(* IEC 61131-3 sources: plc-process-lib/src/POUs/Alarm/FB_Alarm, 9 files *)

(* ---- FB_Alarm.decl.st ---- *)
// Назначение: одна тревога по ISA-18.2. Четыре базовых состояния (Normal, ActiveUnack,
//             ActiveAck, RtnUnack) и три наложенных по старшинству OutOfService >
//             SuppressedByDesign > Shelved; приоритет, задержки появления и снятия (FB_Delay),
//             shelve с таймаутом, подавление по условию, вывод из работы. Каждый переход eState
//             увеличивает udiSeq и отправляет событие в GVL_Lib.itfAlarmSink (если приёмник задан).
//             Методы Ack, Shelve, Unshelve только ставят запрос: его выполняет ближайший вызов тела.
//             Модель состояний и повторное оповещение после shelve — сверить с ANSI/ISA-18.2-2016.
// Автор:      kr0nsch
// Версия:     0.1.0
// Документ:   docs/fb/FB_Alarm.md
FUNCTION_BLOCK FB_Alarm IMPLEMENTS I_Alarm
VAR_INPUT
    xIn           : BOOL;            // условие тревоги (до задержек)
    xSuppress     : BOOL;            // подавление по условию (suppressed by design)
    xOutOfService : BOOL;            // вывод из работы (устройство в OutOfService)
    udiId         : UDINT;           // номер тревоги на объекте
    rValue        : REAL;            // значение процесса для события
    stCfg         : ST_AlarmCfg;     // параметры; 16 байт — копирование дешевле ссылки
    itfTime       : I_TimeSource;    // источник времени; 0 — встроенный fbSysTime
END_VAR
VAR_OUTPUT
    eState        : E_AlarmState := E_AlarmState.Normal;   // состояние ISA-18.2
    xActive       : BOOL;            // условие после задержек (независимо от наложенных состояний)
    xUnacked      : BOOL;            // eState = ActiveUnack OR RtnUnack
    xInList       : BOOL;            // ActiveUnack, ActiveAck или RtnUnack — показывать в списке тревог
    xShelved      : BOOL;            // shelve действует (даже если сверху подавление или OutOfService)
    tShelveRemain : TIME;            // остаток shelve; T#0S — shelve нет
    ltLastChange  : LTIME;           // время последнего перехода
    udiSeq        : UDINT;           // +1 на каждый переход eState (переполнение допустимо)
END_VAR
VAR
    fbDelay      : FB_Delay;         // задержки появления (tOnDelay) и снятия (tOffDelay)
    fbSysTime    : FB_SystemTime;    // запасной источник времени
    xAckReq      : BOOL;             // запрос Ack()
    xShelveReq   : BOOL;             // запрос Shelve()
    tShelveReq   : TIME;             // срок из запроса Shelve()
    xUnshelveReq : BOOL;             // запрос Unshelve()
    ltShelveEnd  : LTIME;            // конец действующего shelve
    // --- реализация (сверх контракта 10.1) ---
    ltNow        : LTIME;            // время этого вызова: отметка переходов и событий
    tShelveDur   : TIME;             // срок действующего shelve (после замены T#0S и обрезки)
    ePrioAct     : E_AlarmPriority := E_AlarmPriority.Medium;      // действующий приоритет
    eShelveEnd   : E_AlarmEventReason := E_AlarmEventReason.None;  // как закончился shelve в этом вызове
END_VAR
VAR_TEMP
    itfTimeAct   : I_TimeSource;     // действующий источник этого вызова
END_VAR

(* ---- FB_Alarm.impl.st ---- *)
// 1. Время этого вызова — один раз, для задержек и для отметок событий
IF itfTime <> 0 THEN
    itfTimeAct := itfTime;
ELSE
    itfTimeAct := fbSysTime;
END_IF
ltNow := itfTimeAct.Now();

// 2. Действующий приоритет: значение вне перечисления (мусор persistent-памяти) считается Medium.
//    Строгое перечисление защищает только исходный текст, поэтому проверка — сравнениями
IF stCfg.ePriority = E_AlarmPriority.None OR stCfg.ePriority = E_AlarmPriority.Low
   OR stCfg.ePriority = E_AlarmPriority.Medium OR stCfg.ePriority = E_AlarmPriority.High
   OR stCfg.ePriority = E_AlarmPriority.Critical
THEN
    ePrioAct := stCfg.ePriority;
ELSE
    ePrioAct := E_AlarmPriority.Medium;
END_IF

IF ePrioAct = E_AlarmPriority.None THEN
    // 3. Тревога выключена: Normal, все выходы FALSE, запросы и shelve снимаются. Если тревога была не в
    //    Normal — один переход с событием Disabled (ALM-1): журнал и сводка по событиям закрывают её; дальше
    //    событий нет. Отсчёт задержки начнётся заново после включения приоритета
    fbDelay.Preset(xValue := FALSE);
    IF eState <> E_AlarmState.Normal THEN
        Transit(eNew := E_AlarmState.Normal, eReason := E_AlarmEventReason.Disabled);
    END_IF
    xActive := FALSE;
    xShelved := FALSE;
    xAckReq := FALSE;
    xShelveReq := FALSE;
    xUnshelveReq := FALSE;
ELSE
    // 4. Условие после задержек появления и снятия
    fbDelay(xIn := xIn, tOnDelay := stCfg.tOnDelay, tOffDelay := stCfg.tOffDelay, itfTime := itfTimeAct);
    xActive := fbDelay.xOut;

    // 5. Квитирование — против состояния на начало вызова; в остальных состояниях без эффекта
    IF xAckReq THEN
        IF eState = E_AlarmState.ActiveUnack THEN
            Transit(eNew := E_AlarmState.ActiveAck, eReason := E_AlarmEventReason.Acked);
        ELSIF eState = E_AlarmState.RtnUnack THEN
            Transit(eNew := E_AlarmState.Normal, eReason := E_AlarmEventReason.Acked);
        END_IF
    END_IF
    xAckReq := FALSE;

    // 6. Shelve: снятие командой, истечение срока, новый запрос
    UpdateShelve();

    // 7–8. Наложенные состояния и базовый автомат ISA-18.2
    UpdateState();
END_IF

// 9. Выходы. После шага 6 при xShelved всегда ltShelveEnd > ltNow: разность без переполнения
xUnacked := eState = E_AlarmState.ActiveUnack OR eState = E_AlarmState.RtnUnack;
xInList := xUnacked OR eState = E_AlarmState.ActiveAck;
IF xShelved THEN
    tShelveRemain := LTIME_TO_TIME(ltShelveEnd - ltNow);
ELSE
    tShelveRemain := T#0S;
END_IF

(* ---- ReleaseState.method.impl.st ---- *)
IF xShelved THEN
    ReleaseState := E_AlarmState.Shelved;
ELSIF xActive THEN
    ReleaseState := E_AlarmState.ActiveUnack;
ELSE
    ReleaseState := E_AlarmState.Normal;
END_IF

(* ---- Shelve.method.decl.st ---- *)
// Запрос shelve; выполняет ближайший вызов тела. TRUE — принято: приоритет не None,
// tShelveMax > 0 и тревога не в OutOfService
METHOD PUBLIC Shelve : BOOL
VAR_INPUT
    tDuration : TIME;   // срок; T#0S — tShelveMax, больше tShelveMax — обрезается
END_VAR

(* ---- Shelve.method.impl.st ---- *)
IF stCfg.ePriority <> E_AlarmPriority.None AND stCfg.tShelveMax > T#0S
   AND eState <> E_AlarmState.OutOfService
THEN
    xShelveReq := TRUE;
    tShelveReq := tDuration;
    Shelve := TRUE;
ELSE
    Shelve := FALSE;
END_IF

(* ---- Transit.method.decl.st ---- *)
// Переход в состояние eNew: udiSeq + 1, отметка времени и событие в GVL_Lib.itfAlarmSink.
// Все переходы ФБ проходят здесь, в порядке шагов тела. Значение процесса в событии всегда конечно:
// NaN и ±Inf (PV из Modbus) — 0.0 (R6). Ответ приёмника (FALSE — переполнен) ФБ
// не повторяет. Внутренний шаг ФБ: PROTECTED, а не PRIVATE (правило L5 контракта)
METHOD PROTECTED Transit
VAR_INPUT
    eNew    : E_AlarmState;          // новое состояние
    eReason : E_AlarmEventReason;    // причина перехода
END_VAR
VAR
    stEvent : ST_AlarmEvent;         // событие для приёмника
END_VAR

(* ---- Transit.method.impl.st ---- *)
stEvent.udiId := udiId;
stEvent.ePriority := ePrioAct;
stEvent.eOldState := eState;
stEvent.eNewState := eNew;
stEvent.eReason := eReason;
stEvent.ltTime := ltNow;
stEvent.rValue := SEL(F_IsFinite(rIn := rValue), 0.0, rValue);

eState := eNew;
udiSeq := udiSeq + 1;
ltLastChange := ltNow;

IF GVL_Lib.itfAlarmSink <> 0 THEN
    GVL_Lib.itfAlarmSink.OnAlarmEvent(stEvent := stEvent);
END_IF

(* ---- UpdateShelve.method.impl.st ---- *)
// 6. Shelve: срок отсчитывается от команды независимо от наложенных состояний
eShelveEnd := E_AlarmEventReason.None;
IF xShelved THEN
    // «время назад»: остаток не может быть больше срока (LTIME без знака — сравнение до вычитания)
    IF ltShelveEnd > ltNow THEN
        IF ltShelveEnd - ltNow > TIME_TO_LTIME(tShelveDur) THEN
            ltShelveEnd := ltNow + TIME_TO_LTIME(tShelveDur);
        END_IF
    END_IF
    IF xUnshelveReq THEN
        xShelved := FALSE;
        eShelveEnd := E_AlarmEventReason.Unshelved;
    ELSIF ltNow >= ltShelveEnd THEN
        xShelved := FALSE;
        eShelveEnd := E_AlarmEventReason.ShelveExpired;
    END_IF
END_IF
// новый запрос (в том числе повторный — срок отсчитывается заново); в OutOfService не принимается
IF xShelveReq AND NOT xOutOfService AND eState <> E_AlarmState.OutOfService
   AND stCfg.tShelveMax > T#0S
THEN
    IF tShelveReq = T#0S OR tShelveReq > stCfg.tShelveMax THEN
        tShelveDur := stCfg.tShelveMax;
    ELSE
        tShelveDur := tShelveReq;
    END_IF
    ltShelveEnd := ltNow + TIME_TO_LTIME(tShelveDur);
    xShelved := TRUE;
    eShelveEnd := E_AlarmEventReason.None;
END_IF
xShelveReq := FALSE;
xUnshelveReq := FALSE;

(* ---- UpdateState.method.impl.st ---- *)
// 7. Наложенные состояния по старшинству OutOfService > SuppressedByDesign > Shelved.
//    Вход — из любого состояния ниже по старшинству (неквитированность сбрасывается),
//    выход — в следующее по старшинству или в базовое: условие активно ? ActiveUnack : Normal
IF xOutOfService THEN
    IF eState <> E_AlarmState.OutOfService THEN
        Transit(eNew := E_AlarmState.OutOfService, eReason := E_AlarmEventReason.OosOn);
    END_IF
ELSIF eState = E_AlarmState.OutOfService THEN
    IF xSuppress THEN
        Transit(eNew := E_AlarmState.SuppressedByDesign, eReason := E_AlarmEventReason.OosOff);
    ELSE
        Transit(eNew := ReleaseState(), eReason := E_AlarmEventReason.OosOff);
    END_IF
ELSIF xSuppress THEN
    IF eState <> E_AlarmState.SuppressedByDesign THEN
        Transit(eNew := E_AlarmState.SuppressedByDesign, eReason := E_AlarmEventReason.Suppressed);
    END_IF
ELSIF eState = E_AlarmState.SuppressedByDesign THEN
    Transit(eNew := ReleaseState(), eReason := E_AlarmEventReason.Unsuppressed);
ELSIF xShelved THEN
    IF eState <> E_AlarmState.Shelved THEN
        Transit(eNew := E_AlarmState.Shelved, eReason := E_AlarmEventReason.Shelved);
    END_IF
ELSIF eState = E_AlarmState.Shelved THEN
    // shelve закончился в этом вызове: командой (Unshelved) или по сроку (ShelveExpired)
    IF eShelveEnd = E_AlarmEventReason.Unshelved THEN
        Transit(eNew := ReleaseState(), eReason := E_AlarmEventReason.Unshelved);
    ELSE
        Transit(eNew := ReleaseState(), eReason := E_AlarmEventReason.ShelveExpired);
    END_IF
// 8. Базовый автомат ISA-18.2
ELSIF eState = E_AlarmState.Normal OR eState = E_AlarmState.RtnUnack THEN
    IF xActive THEN
        Transit(eNew := E_AlarmState.ActiveUnack, eReason := E_AlarmEventReason.Activated);
    END_IF
ELSIF eState = E_AlarmState.ActiveUnack THEN
    IF NOT xActive THEN
        Transit(eNew := E_AlarmState.RtnUnack, eReason := E_AlarmEventReason.Cleared);
    END_IF
ELSIF eState = E_AlarmState.ActiveAck THEN
    IF NOT xActive THEN
        Transit(eNew := E_AlarmState.Normal, eReason := E_AlarmEventReason.Cleared);
    END_IF
END_IF
